Fanuc KAREL source: kd00019.KL

PROGRAM KD00019
%STACKSIZE=65535
%PRIORITY=65535
%NOLOCKGROUP
TYPE
REC_T=STRUCTURE
VALUE : INTEGER
ENDSTRUCTURE
VAR
I : INTEGER
J : INTEGER
B : BOOLEAN
R : REAL
S : STRING[80]
REC : REC_T
BEGIN
REC.VALUE=1
REC.VALUE=(REC.VALUE + 1)
END KD00019
